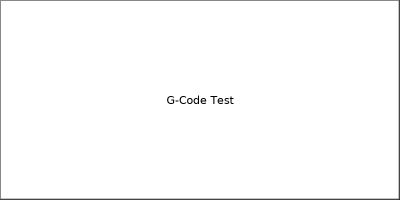
VISUALIZATION V_NCITest  // 400x200
    RoundedRectangle (0,0 400x200)
    Label (93,92 215x17), "G-Code Test"
END_VISUALIZATION

(* stored: Version 1.1.0.1, ProductVersion 3.1.4024.15
   Visu V_NCITest: Id {4a8c3883-2d70-4998-a8f7-7e4f803d03c4} *)
